(* IEC 61131-3 sources: codesys-framework/txt/application/ToDo/Hardware/IO/Cylinder/FB_Cylinder/Properties, 2 files *)

(* ---- State.prop.st ---- *)
PROPERTY State : E_CylinderStates

// --- BEGIN IMPLEMENTATION ---

// ----------- GET -----------
VAR
END_VAR

// -- BEGIN IMPLEMENTATION GET --
State := _eState;

(* ---- SysPar.prop.st ---- *)
PROPERTY SysPar : SC_SystemParametersCylinder

// --- BEGIN IMPLEMENTATION ---

// ----------- SET -----------
VAR
END_VAR

// -- BEGIN IMPLEMENTATION SET --
_scSysPar := SysPar;
